(* IEC 61131-3 sources: llm-plc-st-eval/data/processed_v2/claude-sonnet-4-6/I1/zero_shot, 3 files *)

(* ---- ejec_1.st ---- *)
FUNCTION_BLOCK FB_Semaforo
VAR_INPUT
    habilitado : BOOL; (* Habilita la secuencia normal del semáforo *)
END_VAR

VAR_OUTPUT
    luzV : BOOL; (* Luz verde *)
    luzA : BOOL; (* Luz amarilla *)
    luzR : BOOL; (* Luz roja *)
END_VAR

VAR
    estado      : INT := 0;   (* Estado de la secuencia: 0=Verde, 1=Amarillo, 2=Rojo *)
    timerSec    : TON;        (* Temporizador para la secuencia normal *)
    timerBlink  : TON;        (* Temporizador para el parpadeo de amarillo *)
    blinkOn     : BOOL;       (* Indica si el amarillo intermitente está encendido *)
END_VAR

(* ─────────────────────────────────────────────────────────────────────────── *)
(*  MODO INHABILITADO: amarillo intermitente, verde y rojo apagados            *)
(* ─────────────────────────────────────────────────────────────────────────── *)
IF NOT habilitado THEN

    (* Detener y resetear el temporizador de secuencia *)
    timerSec(IN := FALSE, PT := T#0S);

    (* Resetear estado para que al habilitar de nuevo arranque en verde *)
    estado := 0;

    (* Temporizador de parpadeo: ciclo de 1 segundo *)
    timerBlink(IN := TRUE, PT := T#1S);

    IF timerBlink.Q THEN
        (* Reiniciar el temporizador y alternar el estado del parpadeo *)
        timerBlink(IN := FALSE, PT := T#1S);
        blinkOn := NOT blinkOn;
    END_IF;

    (* Asignar salidas: solo amarillo parpadea *)
    luzV := FALSE;
    luzA := blinkOn;
    luzR := FALSE;

(* ─────────────────────────────────────────────────────────────────────────── *)
(*  MODO HABILITADO: secuencia Verde → Amarillo → Rojo                        *)
(* ─────────────────────────────────────────────────────────────────────────── *)
ELSE

    (* Detener y resetear el temporizador de parpadeo *)
    timerBlink(IN := FALSE, PT := T#0S);
    blinkOn := FALSE;

    CASE estado OF

        (* ── Estado 0: Verde 20 s ── *)
        0:
            luzV := TRUE;
            luzA := FALSE;
            luzR := FALSE;

            timerSec(IN := TRUE, PT := T#20S);
            IF timerSec.Q THEN
                timerSec(IN := FALSE, PT := T#20S); (* Resetear temporizador *)
                estado := 1;                         (* Pasar a amarillo *)
            END_IF;

        (* ── Estado 1: Amarillo 4 s ── *)
        1:
            luzV := FALSE;
            luzA := TRUE;
            luzR := FALSE;

            timerSec(IN := TRUE, PT := T#4S);
            IF timerSec.Q THEN
                timerSec(IN := FALSE, PT := T#4S);  (* Resetear temporizador *)
                estado := 2;                         (* Pasar a rojo *)
            END_IF;

        (* ── Estado 2: Rojo 15 s ── *)
        2:
            luzV := FALSE;
            luzA := FALSE;
            luzR := TRUE;

            timerSec(IN := TRUE, PT := T#15S);
            IF timerSec.Q THEN
                timerSec(IN := FALSE, PT := T#15S); (* Resetear temporizador *)
                estado := 0;                         (* Volver a verde *)
            END_IF;

        (* ── Estado por defecto: seguridad ── *)
        ELSE
            estado := 0;
            timerSec(IN := FALSE, PT := T#0S);

    END_CASE;

END_IF;

(* ---- ejec_2.st ---- *)
FUNCTION_BLOCK FB_Semaforo
VAR_INPUT
    habilitado : BOOL; (* Habilita la secuencia normal del semáforo *)
END_VAR

VAR_OUTPUT
    luzV : BOOL; (* Luz verde *)
    luzA : BOOL; (* Luz amarilla *)
    luzR : BOOL; (* Luz roja *)
END_VAR

VAR
    (* Temporizadores TON estándar IEC 61131-3 *)
    tVerde      : TON; (* Temporiza la fase verde  - 20 s *)
    tAmarillo   : TON; (* Temporiza la fase amarilla - 4 s *)
    tRojo       : TON; (* Temporiza la fase roja   - 15 s *)
    tParpadeo   : TON; (* Temporiza el parpadeo amarillo - 1 s *)

    (* Estado de la secuencia normal *)
    (* 0 = Verde, 1 = Amarillo, 2 = Rojo *)
    estado      : INT := 0;

    (* Bit de parpadeo para amarillo intermitente *)
    parpadeo    : BOOL := FALSE;
END_VAR

(* ─────────────────────────────────────────────────────────────
   MODO DESHABILITADO: amarillo intermitente, resto apagado
   ───────────────────────────────────────────────────────────── *)
IF NOT habilitado THEN

    (* Reiniciar estado para que al habilitar arranque en verde *)
    estado := 0;

    (* Apagar temporizadores de secuencia normal *)
    tVerde(IN := FALSE,   PT := T#20S);
    tAmarillo(IN := FALSE, PT := T#4S);
    tRojo(IN := FALSE,    PT := T#15S);

    (* Temporizador de parpadeo: ciclo de 1 s *)
    tParpadeo(IN := TRUE, PT := T#1S);

    IF tParpadeo.Q THEN
        (* Reiniciar temporizador y conmutar estado de parpadeo *)
        tParpadeo(IN := FALSE, PT := T#1S);
        parpadeo := NOT parpadeo;
    END_IF;

    (* Salidas: solo amarillo parpadea *)
    luzV := FALSE;
    luzA := parpadeo;
    luzR := FALSE;

(* ─────────────────────────────────────────────────────────────
   MODO HABILITADO: secuencia Verde → Amarillo → Rojo → ...
   ───────────────────────────────────────────────────────────── *)
ELSE

    (* Detener temporizador de parpadeo y resetear bit *)
    tParpadeo(IN := FALSE, PT := T#1S);
    parpadeo := FALSE;

    CASE estado OF

        (* ── FASE VERDE ── *)
        0:
            luzV := TRUE;
            luzA := FALSE;
            luzR := FALSE;

            tVerde(IN := TRUE, PT := T#20S);

            IF tVerde.Q THEN
                (* Verde cumplido → pasar a amarillo *)
                tVerde(IN := FALSE, PT := T#20S); (* Reset temporizador *)
                estado := 1;
            END_IF;

        (* ── FASE AMARILLO ── *)
        1:
            luzV := FALSE;
            luzA := TRUE;
            luzR := FALSE;

            tAmarillo(IN := TRUE, PT := T#4S);

            IF tAmarillo.Q THEN
                (* Amarillo cumplido → pasar a rojo *)
                tAmarillo(IN := FALSE, PT := T#4S); (* Reset temporizador *)
                estado := 2;
            END_IF;

        (* ── FASE ROJO ── *)
        2:
            luzV := FALSE;
            luzA := FALSE;
            luzR := TRUE;

            tRojo(IN := TRUE, PT := T#15S);

            IF tRojo.Q THEN
                (* Rojo cumplido → volver a verde *)
                tRojo(IN := FALSE, PT := T#15S); (* Reset temporizador *)
                estado := 0;
            END_IF;

        (* ── ESTADO INVÁLIDO: recuperar a verde ── *)
        ELSE
            estado := 0;

    END_CASE;

END_IF;

(* ---- ejec_3.st ---- *)
FUNCTION_BLOCK FB_Semaforo
VAR_INPUT
    habilitado : BOOL; (* Habilita la secuencia normal del semáforo *)
END_VAR

VAR_OUTPUT
    luzV : BOOL; (* Luz verde *)
    luzA : BOOL; (* Luz amarilla *)
    luzR : BOOL; (* Luz roja *)
END_VAR

VAR
    (* Temporizadores TON estándar IEC 61131-3 *)
    tVerde      : TON; (* Temporizador fase verde  - 20 s *)
    tAmarillo   : TON; (* Temporizador fase amarilla - 4 s *)
    tRojo       : TON; (* Temporizador fase roja   - 15 s *)
    tParpadeo   : TON; (* Temporizador parpadeo amarillo - 1 s *)

    (* Estado interno de la secuencia normal *)
    (* 0 = Verde, 1 = Amarillo, 2 = Rojo *)
    estado      : INT := 0;

    (* Bit de parpadeo para amarillo intermitente *)
    bitParpadeo : BOOL := FALSE;
END_VAR

(* ─────────────────────────────────────────────────────────────
   MODO INHABILITADO: amarillo intermitente, resto apagado
   ───────────────────────────────────────────────────────────── *)
IF NOT habilitado THEN

    (* Reiniciar la secuencia para que arranque en verde al volver *)
    estado := 0;

    (* Apagar temporizadores de secuencia normal *)
    tVerde(IN := FALSE,    PT := T#20S);
    tAmarillo(IN := FALSE, PT := T#4S);
    tRojo(IN := FALSE,     PT := T#15S);

    (* Parpadeo: el temporizador cuenta 1 s; al vencer, invierte el bit *)
    tParpadeo(IN := TRUE, PT := T#1S);
    IF tParpadeo.Q THEN
        bitParpadeo := NOT bitParpadeo;
        tParpadeo(IN := FALSE, PT := T#1S); (* Reinicia el temporizador *)
    END_IF;

    (* Salidas: solo amarillo parpadea *)
    luzV := FALSE;
    luzA := bitParpadeo;
    luzR := FALSE;

(* ─────────────────────────────────────────────────────────────
   MODO HABILITADO: secuencia Verde → Amarillo → Rojo → ...
   ───────────────────────────────────────────────────────────── *)
ELSE

    (* Detener temporizador de parpadeo y resetear bit *)
    tParpadeo(IN := FALSE, PT := T#1S);
    bitParpadeo := FALSE;

    CASE estado OF

        (* ── FASE VERDE (20 s) ── *)
        0:
            luzV := TRUE;
            luzA := FALSE;
            luzR := FALSE;

            tVerde(IN := TRUE, PT := T#20S);
            IF tVerde.Q THEN
                tVerde(IN := FALSE, PT := T#20S); (* Reinicia temporizador *)
                estado := 1;                       (* Pasa a amarillo *)
            END_IF;

        (* ── FASE AMARILLO (4 s) ── *)
        1:
            luzV := FALSE;
            luzA := TRUE;
            luzR := FALSE;

            tAmarillo(IN := TRUE, PT := T#4S);
            IF tAmarillo.Q THEN
                tAmarillo(IN := FALSE, PT := T#4S); (* Reinicia temporizador *)
                estado := 2;                         (* Pasa a rojo *)
            END_IF;

        (* ── FASE ROJO (15 s) ── *)
        2:
            luzV := FALSE;
            luzA := FALSE;
            luzR := TRUE;

            tRojo(IN := TRUE, PT := T#15S);
            IF tRojo.Q THEN
                tRojo(IN := FALSE, PT := T#15S); (* Reinicia temporizador *)
                estado := 0;                      (* Vuelve a verde *)
            END_IF;

        (* ── ESTADO INVÁLIDO: recuperación segura ── *)
        ELSE
            estado := 0;
            luzV := FALSE;
            luzA := FALSE;
            luzR := FALSE;

    END_CASE;

END_IF;

END_FUNCTION_BLOCK
